{attribute 'qualified_only'}
{attribute 'strict'}
{attribute 'to_string'}
TYPE EN_Pump_SPAL_ServiceIndicator :
(
   Not_Available,
   Reserved,
   Service_required,
   Service_not_required
);
END_TYPE

(* stored: Version 1.1.0.1
   DUT EN_Pump_SPAL_ServiceIndicator: Id {fe68fd77-9c9b-4194-8e90-56313d8b294a} *)
